// TwinCAT 3 PLC project Untitled1
// ProgramVersion: 3.1.4026.25
// libraries:
//   Tc2_Standard, * (Beckhoff Automation GmbH)
//   Tc2_System, * (Beckhoff Automation GmbH)
// project tree:
//   GVLs/ GVL_Inputs.TcGVL, GVL_IO.TcGVL, GVL_Outputs.TcGVL
//   / PlcTask.TcTTO
//   POUs/ MAIN.TcPOU, PRG_Mapping.TcPOU
// real-time tasks:
//   TASK PlcTask: cycle T#10ms, priority 20, ADS port 350
// I/O:
//   DEVICE Device 1 (EtherCAT), AmsNetId 192.168.0.210.2.1
//     +MP-5K1 (CU1128) [CU1128 6x EtherCAT junction]
//       +MP-6K1(EK1100) [EK1100 EtherCAT Coupler (2A E-Bus)]
//         +MP-6K10(EL1809) [EL1809 16Ch. Dig. Input 24V, 3ms]
//         +MP-6K20(EL2809) [EL2809 16Ch. Dig. Output 24V, 0.5A]
//         Analog input (EL3102) [EL3102 2Ch. Ana. Input +/-10V, Diff.]
//         Temp Sensor (EL3204) [EL3204 4Ch. Ana. Input PT100 (RTD)]
//         Encoder (EL5101) [EL5101 1Ch. Inc. Encoder 5V]
//       Box 2 (CU1128-B) [CU1128 6x EtherCAT junction - Dev A]
//         +LS-7K1 (EK1100) [EK1100 EtherCAT Coupler (2A E-Bus)]
//           Term 8 (EL1809) [EL1809 16Ch. Dig. Input 24V, 3ms]
//           Term 9 (EL2809) [EL2809 16Ch. Dig. Output 24V, 0.5A]
//       Box 3 (CU1128-C) [CU1128 6x EtherCAT junction - Dev B]
//         +MS-9K1 (EP1018-0001) [EP1018-0001 8 Ch. Dig. Input 24V, 10µs, M8]
//         +MS-9K2 (EP1018-0001) [EP1018-0001 8 Ch. Dig. Input 24V, 10µs, M8]
//         +MS-9K3 (EP1018-0001) [EP1018-0001 8 Ch. Dig. Input 24V, 10µs, M8]
//         +MS-10K1 (EP2028-0001) [EP2028-0001 8 Ch. Dig. Output 24V, 2A, M8]
//         +MS-10K2 (EP2028-0001) [EP2028-0001 8 Ch. Dig. Output 24V, 2A, M8]

CONFIGURATION Untitled1
    RESOURCE PLC ON TwinCAT3
        TASK PlcTask(INTERVAL := T#10ms, PRIORITY := 20);
        PROGRAM MAIN WITH PlcTask : MAIN;
    END_RESOURCE
END_CONFIGURATION

// ---- GVLs/GVL_Inputs.TcGVL
{attribute 'qualified_only'}
VAR_GLOBAL

    // === INPUTS: MAIN CONTROL CABINET & SPECIAL MODULES ==================

    bAirServiceUnit_PressureOK  : BOOL;  // Main Cabinet Pressure Switch
    bEStop_Pressed              : BOOL;  // Main Cabinet Emergency Stop
    
    nAnalog_Pressure_Sensor     : INT;   // EL3102 Analog Value
    nTemp_Heater_Band           : INT;   // EL3204 Temp Value
    
    nEncoder_Position           : UDINT; // EL5101 Counter Value
    bEncoder_Latch              : BOOL;  // EL5101 Status Latch


    // === INPUTS: SECONDARY STATION / LASER SYSTEM ========================

    bCW_Ready                   : BOOL;
    bCW_AckCoded                : BOOL;
    bCW_MarkInProgress          : BOOL;

    // === INPUTS: DECENTRALIZED FIELD BOXES (Cylinder & Sensor states) ====
    
    // Box 1
    bCyl_Ejector_Ext            : BOOL;  
    bCyl_Ejector_Ret            : BOOL;  
    bCyl_Clamp_Ext              : BOOL;  
    bCyl_Clamp_Ret              : BOOL;  
    bCyl_Diverter_Ext           : BOOL;  
    bCyl_Diverter_Ret           : BOOL;  

    // Box 2
    bCyl_Infeed_Ext             : BOOL;  
    bCyl_Infeed_Ret             : BOOL;  
    bCyl_Outfeed_Ext            : BOOL;  
    bCyl_Outfeed_Ret            : BOOL;  

    // Box 3
    bLightBarrier_Infeed        : BOOL;  
    bServo_Infeed_Locked        : BOOL;  
    bServo_Infeed_AS            : BOOL;  
    bServo_Infeed_GS            : BOOL;  
    bLightBarrier_Outfeed       : BOOL;  
    bServo_Outfeed_Locked       : BOOL;  
    bServo_Outfeed_AS           : BOOL;  
    bServo_Outfeed_GS           : BOOL;

END_VAR

// ---- GVLs/GVL_IO.TcGVL
{attribute 'qualified_only'}
VAR_GLOBAL
		// --- Digital Inputs (Term 5: EL1809) ---
    bAirServiceUnit_PressureOK  AT %I* : BOOL;  // EL1809 Ch 1 (Pressure switch +MS-12B1)
    bEStop_Pressed              AT %I* : BOOL;  // EL1809 Ch 2 (Emergency Stop +BP1-8S1)
    
    // --- Digital Outputs (Term 6: EL2809) ---
    bAirServiceUnit_Vent        AT %Q* : BOOL;  // EL2809 Ch 1 (Vent valve +MS-12Q1)
    bLaserEnable                AT %Q* : BOOL;  // EL2809 Ch 2 (Laser Enable Relay)
    
    // --- Analog Inputs (EL3102) ---
    nAnalog_Pressure_Sensor     AT %I* : INT;   // EL3102 Ch 1 (0-10V or 4-20mA raw value)
    
    // --- Temperature Measurement (EL3204) ---
    nTemp_Heater_Band           AT %I* : INT;   // EL3204 Ch 1 (PT100 temperature value)
    
    // --- Counter / Encoder Module (EL5101) ---
    nEncoder_Position           AT %I* : UDINT; // EL5101 Counter Value
    bEncoder_Latch              AT %I* : BOOL;  // EL5101 Status / Latch
    
    // --- CW Controller Inputs (EL1809) ---
    bCW_Ready                   AT %I* : BOOL;  // Secondary EL1809 Ch 1
    bCW_AckCoded                AT %I* : BOOL;  // Secondary EL1809 Ch 2
    bCW_MarkInProgress          AT %I* : BOOL;  // Secondary EL1809 Ch 3
    
    // --- CW Controller Outputs (EL2809) ---
    bCW_DWTrig                  AT %Q* : BOOL;  // Secondary EL2809 Ch 1

    // --- Field Input Box 1: +MS-9K1 (EP1018-0001) ---
    bCyl_Ejector_Ext            AT %I* : BOOL;  // EP1018 Box 1 Ch 1
    bCyl_Ejector_Ret            AT %I* : BOOL;  // EP1018 Box 1 Ch 2 
    bCyl_Clamp_Ext              AT %I* : BOOL;  // EP1018 Box 1 Ch 3
    bCyl_Clamp_Ret              AT %I* : BOOL;  // EP1018 Box 1 Ch 4 
    bCyl_Diverter_Ext           AT %I* : BOOL;  // EP1018 Box 1 Ch 5 
    bCyl_Diverter_Ret           AT %I* : BOOL;  // EP1018 Box 1 Ch 6 

    // --- Field Input Box 2: +MS-9K2 (EP1018-0001) ---
    bCyl_Infeed_Ext             AT %I* : BOOL;  // EP1018 Box 2 Ch 1 
    bCyl_Infeed_Ret             AT %I* : BOOL;  // EP1018 Box 2 Ch 2 
    bCyl_Outfeed_Ext            AT %I* : BOOL;  // EP1018 Box 2 Ch 3 
    bCyl_Outfeed_Ret            AT %I* : BOOL;  // EP1018 Box 2 Ch 4 

    // --- Field Input Box 3: +MS-9K3 (EP1018-0001) ---
    bLightBarrier_Infeed        AT %I* : BOOL;  // EP1018 Box 3 Ch 1 
    bServo_Infeed_Locked        AT %I* : BOOL;  // EP1018 Box 3 Ch 2 
    bServo_Infeed_AS            AT %I* : BOOL;  // EP1018 Box 3 Ch 3 
    bServo_Infeed_GS            AT %I* : BOOL;  // EP1018 Box 3 Ch 4 
    bLightBarrier_Outfeed       AT %I* : BOOL;  // EP1018 Box 3 Ch 5 
    bServo_Outfeed_Locked       AT %I* : BOOL;  // EP1018 Box 3 Ch 6 
    bServo_Outfeed_AS           AT %I* : BOOL;  // EP1018 Box 3 Ch 7 
    bServo_Outfeed_GS           AT %I* : BOOL;  // EP1018 Box 3 Ch 8
    
    // --- Field Output Box 1: +MS-10K1 (EP2028-0001) ---
    bValve_Ejector_Ext          AT %Q* : BOOL;  // EP2028 Box 1 Ch 1 
    bValve_Ejector_Ret          AT %Q* : BOOL;  // EP2028 Box 1 Ch 2 
    bValve_Clamp_Ext            AT %Q* : BOOL;  // EP2028 Box 1 Ch 3 
    bValve_Clamp_Ret            AT %Q* : BOOL;  // EP2028 Box 1 Ch 4 
    bValve_Diverter_Ext         AT %Q* : BOOL;  // EP2028 Box 1 Ch 5 
    bValve_Diverter_Ret         AT %Q* : BOOL;  // EP2028 Box 1 Ch 6 

    // --- Field Output Box 2: +MS-10K2 (EP2028-0001) ---
    bValve_Infeed_Ext           AT %Q* : BOOL;  // EP2028 Box 2 Ch 1 
    bValve_Infeed_Ret           AT %Q* : BOOL;  // EP2028 Box 2 Ch 2 
    bValve_Outfeed_Ext          AT %Q* : BOOL;  // EP2028 Box 2 Ch 3 
    bValve_Outfeed_Ret          AT %Q* : BOOL;  // EP2028 Box 2 Ch 4 
    bValve_AirBlow_AS           AT %Q* : BOOL;  // EP2028 Box 2 Ch 5 
    bValve_AirBlow_GS           AT %Q* : BOOL;  // EP2028 Box 2 Ch 6 
    bValve_Bypass_AS            AT %Q* : BOOL;  // EP2028 Box 2 Ch 7 
    bValve_Bypass_GS            AT %Q* : BOOL;  // EP2028 Box 2 Ch 8 
END_VAR

// ---- GVLs/GVL_Outputs.TcGVL
{attribute 'qualified_only'}
VAR_GLOBAL

    // === OUTPUTS: MAIN CONTROL CABINET & LASER SYSTEM ====================

    bAirServiceUnit_Vent        : BOOL;  // Main Cabinet Vent Valve
    bLaserEnable                : BOOL;  // Main Cabinet Laser Enable Relay
    
    bCW_DWTrig                  : BOOL;  // Laser System Trigger

    // === OUTPUTS: DECENTRALIZED FIELD BOXES (Pneumatic Valves) ===========

    // Box 1
    bValve_Ejector_Ext          : BOOL;  
    bValve_Ejector_Ret          : BOOL;  
    bValve_Clamp_Ext            : BOOL;  
    bValve_Clamp_Ret            : BOOL;  
    bValve_Diverter_Ext         : BOOL;  
    bValve_Diverter_Ret         : BOOL;  

    // Box 2
    bValve_Infeed_Ext           : BOOL;  
    bValve_Infeed_Ret           : BOOL;  
    bValve_Outfeed_Ext          : BOOL;  
    bValve_Outfeed_Ret          : BOOL;  
    bValve_AirBlow_AS           : BOOL;  
    bValve_AirBlow_GS           : BOOL;  
    bValve_Bypass_AS            : BOOL;  
    bValve_Bypass_GS            : BOOL;
END_VAR

// ---- POUs/MAIN.TcPOU
PROGRAM MAIN
VAR
END_VAR

// Call I/O Mapping Program
PRG_Mapping();

END_PROGRAM

// ---- POUs/PRG_Mapping.TcPOU
PROGRAM PRG_Mapping
VAR
END_VAR


// === READ INPUTS (Hardware -> Software) ==============================

// --- Main Control Cabinet & Special Modules ---
GVL_Inputs.bAirServiceUnit_PressureOK := GVL_IO.bAirServiceUnit_PressureOK;
GVL_Inputs.bEStop_Pressed             := GVL_IO.bEStop_Pressed;
GVL_Inputs.nAnalog_Pressure_Sensor    := GVL_IO.nAnalog_Pressure_Sensor;
GVL_Inputs.nTemp_Heater_Band          := GVL_IO.nTemp_Heater_Band;
GVL_Inputs.nEncoder_Position          := GVL_IO.nEncoder_Position;
GVL_Inputs.bEncoder_Latch             := GVL_IO.bEncoder_Latch;

// --- Secondary Station / Laser System ---
GVL_Inputs.bCW_Ready                  := GVL_IO.bCW_Ready;
GVL_Inputs.bCW_AckCoded               := GVL_IO.bCW_AckCoded;
GVL_Inputs.bCW_MarkInProgress         := GVL_IO.bCW_MarkInProgress;

// --- Decentralized Field Box 1 ---
GVL_Inputs.bCyl_Ejector_Ext           := GVL_IO.bCyl_Ejector_Ext;
GVL_Inputs.bCyl_Ejector_Ret           := GVL_IO.bCyl_Ejector_Ret;
GVL_Inputs.bCyl_Clamp_Ext             := GVL_IO.bCyl_Clamp_Ext;
GVL_Inputs.bCyl_Clamp_Ret             := GVL_IO.bCyl_Clamp_Ret;
GVL_Inputs.bCyl_Diverter_Ext          := GVL_IO.bCyl_Diverter_Ext;
GVL_Inputs.bCyl_Diverter_Ret          := GVL_IO.bCyl_Diverter_Ret;

// --- Decentralized Field Box 2 ---
GVL_Inputs.bCyl_Infeed_Ext            := GVL_IO.bCyl_Infeed_Ext;
GVL_Inputs.bCyl_Infeed_Ret            := GVL_IO.bCyl_Infeed_Ret;
GVL_Inputs.bCyl_Outfeed_Ext           := GVL_IO.bCyl_Outfeed_Ext;
GVL_Inputs.bCyl_Outfeed_Ret           := GVL_IO.bCyl_Outfeed_Ret;

// --- Decentralized Field Box 3 ---
GVL_Inputs.bLightBarrier_Infeed       := GVL_IO.bLightBarrier_Infeed;
GVL_Inputs.bServo_Infeed_Locked       := GVL_IO.bServo_Infeed_Locked;
GVL_Inputs.bServo_Infeed_AS           := GVL_IO.bServo_Infeed_AS;
GVL_Inputs.bServo_Infeed_GS           := GVL_IO.bServo_Infeed_GS;
GVL_Inputs.bLightBarrier_Outfeed      := GVL_IO.bLightBarrier_Outfeed;
GVL_Inputs.bServo_Outfeed_Locked      := GVL_IO.bServo_Outfeed_Locked;
GVL_Inputs.bServo_Outfeed_AS          := GVL_IO.bServo_Outfeed_AS;
GVL_Inputs.bServo_Outfeed_GS          := GVL_IO.bServo_Outfeed_GS;

// === WRITE OUTPUTS (Software -> Hardware) ============================

// --- Main Control Cabinet & Laser System ---
GVL_IO.bAirServiceUnit_Vent           := GVL_Outputs.bAirServiceUnit_Vent;
GVL_IO.bLaserEnable                   := GVL_Outputs.bLaserEnable;
GVL_IO.bCW_DWTrig                     := GVL_Outputs.bCW_DWTrig;

// --- Decentralized Field Box 1 ---
GVL_IO.bValve_Ejector_Ext             := GVL_Outputs.bValve_Ejector_Ext;
GVL_IO.bValve_Ejector_Ret             := GVL_Outputs.bValve_Ejector_Ret;
GVL_IO.bValve_Clamp_Ext               := GVL_Outputs.bValve_Clamp_Ext;
GVL_IO.bValve_Clamp_Ret               := GVL_Outputs.bValve_Clamp_Ret;
GVL_IO.bValve_Diverter_Ext            := GVL_Outputs.bValve_Diverter_Ext;
GVL_IO.bValve_Diverter_Ret            := GVL_Outputs.bValve_Diverter_Ret;

// --- Decentralized Field Box 2 ---
GVL_IO.bValve_Infeed_Ext              := GVL_Outputs.bValve_Infeed_Ext;
GVL_IO.bValve_Infeed_Ret              := GVL_Outputs.bValve_Infeed_Ret;
GVL_IO.bValve_Outfeed_Ext             := GVL_Outputs.bValve_Outfeed_Ext;
GVL_IO.bValve_Outfeed_Ret             := GVL_Outputs.bValve_Outfeed_Ret;
GVL_IO.bValve_AirBlow_AS              := GVL_Outputs.bValve_AirBlow_AS;
GVL_IO.bValve_AirBlow_GS              := GVL_Outputs.bValve_AirBlow_GS;
GVL_IO.bValve_Bypass_AS               := GVL_Outputs.bValve_Bypass_AS;
GVL_IO.bValve_Bypass_GS               := GVL_Outputs.bValve_Bypass_GS;

END_PROGRAM
